// TIA Portal V20 export
// export: Created 2026-10-12T05:35:24.8995057Z, ExportSetting WithDefaults, DisplayName Totally Integrated Automation Portal, DisplayVersion V20, DisplayName TIA Portal Openness, DisplayVersion V20, DisplayName TIA Portal Teamcenter Gateway, DisplayVersion V20, DisplayName TIA Portal Version Control Interface, DisplayVersion V20, DisplayName SINAMICS Startdrive Advanced, DisplayVersion V20 SP1 Update 2, DisplayName SINAMICS Startdrive G110M, G120, G120C, G120D, G120P, G115D, DisplayVersion V20 SP1 Update 2, DisplayName SINAMICS Startdrive G130, G150, S120, S150, SINAMICS MV, G220, S200, S210, DisplayVersion V20 SP1 Update 2, DisplayName STEP 7 Professional, DisplayVersion V20, DisplayName STEP 7 Safety, DisplayVersion V20, DisplayName WinCC Basic/Comfort/Advanced, DisplayVersion V20, DisplayName WinCC Professional, DisplayVersion V20, DisplayName WinCC Unified, DisplayVersion V20
FUNCTION "FRK_PathOwned" : Bool   // FC79, SCL
{ S7_Optimized_Access := 'TRUE' }
VERSION : 0.1
// Shared Unit routing: typed generated edges carry these owning predicates.
// stored: AutoNumber true, IsIECCheckEnabled false, SetENOAutomatically false, UDAEnableTagReadback false
   VAR_INPUT
      OwnerPath : String;
      TargetPath : WString;
   END_VAR
   VAR_TEMP
      Width : Int;
   END_VAR
BEGIN

   #FRK_PathOwned := FALSE;
   #Width := LEN(#OwnerPath);
   IF #Width = 0 THEN
       RETURN;
   END_IF;
   IF #TargetPath = STRING_TO_WSTRING(#OwnerPath) THEN
       #FRK_PathOwned := TRUE;
       RETURN;
   END_IF;
   IF LEN(#TargetPath) <= #Width THEN
       RETURN;
   END_IF;
   #FRK_PathOwned := LEFT(IN := #TargetPath, L := #Width) = STRING_TO_WSTRING(#OwnerPath) AND #TargetPath[#Width + 1] = WCHAR#'.';
END_FUNCTION
